TYPE ST_EntrywayInputs :
STRUCT
    bLowerButton : BOOL;
    bUpperButton : BOOL;
END_STRUCT
END_TYPE

(* stored: Version 1.1.0.1
   DUT ST_EntrywayInputs: Id {c7580358-4cba-4ea5-a8b1-488aab250f69} *)
